(* IEC 61131-3 sources: Codesys_IAP/Demo/PLC1/PLC 1 Simulatie Ladder StructuredTekst IOStructures 2V0_tekst/Programma Structured Text/Structures, 7 files *)

(* ---- hmiIO.st ---- *)
(*#### DECLARATIE ####*)
// Datum : 17 december 2020, Auteur: Gerard Harkema
TYPE hmiIO :
STRUCT
	// Indrukken resetknop
	Ix_Resetknop			: REFERENCE TO BOOL;
	// Keuzeknop staat op hand
	Ix_Hand					: REFERENCE TO BOOL;
	// Keuzeknop staat op auto
	Ix_Auto					: REFERENCE TO BOOL;
	// Indrukken noodstop
	Ix_Noodstop				: REFERENCE TO BOOL;
	// Bekers magazijn zijn op

	// Indrukken startknop
	Ix_Stopknop				: REFERENCE TO BOOL;
	// Indrukken stopknop
	Ix_Startknop			: REFERENCE TO BOOL;
	//Perslucht is aanwezig

	// Visualisatie invisible Gele vlak
	Qx_GeleLamp				: REFERENCE TO BOOL;
	// Visualisatie invisible groene vlak
	Qx_GroeneLamp			: REFERENCE TO BOOL;
	// Visualisatie invisible rode vlak
	Qx_RodeLamp				: REFERENCE TO BOOL;

END_STRUCT
END_TYPE

(* ---- magazijnIO.st ---- *)
(*#### DECLARATIE ####*)
// Datum : 17 december 2020, Auteur: Gerard Harkema
TYPE magazijnIO :
STRUCT
	// Bekers magazijn zijn op
	Ix_MagazijnLeeg				: REFERENCE TO BOOL;
	// Beker is uit dekselmagazijn gestoten
	Ix_UitstoterBekerIn			: REFERENCE TO BOOL;
	// Uitstoter Beker haalt nieuwe beker op
	Ix_UitstoterBekerUit		: REFERENCE TO BOOL;
	// Beker uit magazijn stoten
	Qx_BekerUitstoten			: REFERENCE TO BOOL;

	//Perslucht is aanwezig
	Ix_PersluchtAanwezig 		: REFERENCE TO BOOL;

END_STRUCT
END_TYPE

(* ---- meetstationIO.st ---- *)
(*#### DECLARATIE ####*)
// Datum : 17 december 2020, Auteur: Gerard Harkema
TYPE meetstationIO :
STRUCT
	//Beker aanwezig op detectiepositie
	Ix_BekerAanwezig :REFERENCE TO BOOL;
	//Beker is van aluminium
	Ix_BekerMetaal :REFERENCE TO BOOL;
	//Beker reflecteert en is dus niet zwart
	Ix_BekerReflecteerd :REFERENCE TO BOOL;
END_STRUCT
END_TYPE

(* ---- overzetterIO.st ---- *)
(*#### DECLARATIE ####*)
// Datum : 17 december 2020, Auteur: Gerard Harkema
TYPE overzetterIO :
STRUCT
	//Werkstuk door overzetter opgepakt
	Ix_VacuumAanwezig 		:REFERENCE TO BOOL;
	//Overzetter haalt beker op(linker pos.)
	Ix_OverzetterIsLinks 	:REFERENCE TO BOOL;
	//Overzetter plaatst beker op sorteerpositie
	Ix_OverzetterIsRechts 	:REFERENCE TO BOOL;
	//Beker aanwezig op detectiepositie

		//Beker oppakken
	Qx_VacuumAan 			:REFERENCE TO BOOL;
	//Beker loslaten
	Qx_BekerLossen 			:REFERENCE TO BOOL;
	//Overzetter naar bekermagazijn
	Qx_OverzetterLinks 		:REFERENCE TO BOOL;
	//Overzetter naar sorteerpositie
	Qx_OverzetterRechts 	:REFERENCE TO BOOL;

END_STRUCT
END_TYPE

(* ---- sorteerGootIO.st ---- *)
(*#### DECLARATIE ####*)
// Datum : 17 december 2020, Auteur: Gerard Harkema
TYPE sorteerGootIO :
STRUCT
		//Product is naar een van de goten gegaan
	Ix_BekerInGoot 			:REFERENCE TO BOOL;
	//Pusher uitvoergoot 1 is in
	Ix_UitvoerGoot1IsIn 	:REFERENCE TO BOOL;
	//Pusher uitvoergoot 2 is in
	Ix_UitvoerGoot2IsIn 	:REFERENCE TO BOOL;
	//Pusher uitvoergoot 3 is in
	Ix_UitvoerGoot3IsIn 	:REFERENCE TO BOOL;
	//Beker afvoeren is bezig
	Ix_StationAfvoerVrij 	:REFERENCE TO BOOL;
	//Pusher uitvoergoot 1 is uit
	Ix_UitvoerGoot1IsUit 	:REFERENCE TO BOOL;
	//Pusher uitvoergoot 2 is uit
	Ix_UitvoerGoot2IsUit 	:REFERENCE TO BOOL;
	//Pusher uitvoergoot 3 is uit
	Ix_UitvoerGoot3IsUit 	:REFERENCE TO BOOL;

	//Transportband aan
	Qx_MotorAfvoerAan 		:REFERENCE TO BOOL;
	//Pusher goot 1 uit
	Qx_UitvoerGoot1Uit 		:REFERENCE TO BOOL;
	//Pusher goot 2 uit
	Qx_UitvoerGoot2Uit 		:REFERENCE TO BOOL;
	//Pusher goot 3 uit
	Qx_UitvoerGoot3Uit 		:REFERENCE TO BOOL;
	//Beker stoppen op band voor detectie
	Qx_StopperUit 			:REFERENCE TO BOOL;
	//Uitsorteren is bezet
	Qx_StationBezet 		:REFERENCE TO BOOL;

	uitvoerGoot1			:uitvoerGootIO;
	uitvoerGoot2			:uitvoerGootIO;
	uitvoerGoot3			:uitvoerGootIO;
	meetstation				:meetstationIO;

END_STRUCT
END_TYPE

(* ---- sorteerStationIO.st ---- *)
(*#### DECLARATIE ####*)
// Datum : 17 december 2020, Auteur: Gerard Harkema
TYPE sorteerStationIO :
STRUCT
	magazijn		: magazijnIO;
	overzetter		: overzetterIO;
	sorteerGoot		: sorteerGootIO;
	hmi				: hmiIO;
END_STRUCT
END_TYPE

(* ---- uitvoerGootIO.st ---- *)
(*#### DECLARATIE ####*)
// Datum : 17 december 2020, Auteur: Gerard Harkema
TYPE uitvoerGootIO :
STRUCT
	//Pusher uitvoergoo is in
	Ix_UitvoerGootIsIn 		: REFERENCE TO BOOL;
	//Pusher uitvoergoot is uit
	Ix_UitvoerGootIsUit 	: REFERENCE TO BOOL;
	//Pusher goot uit
	Qx_UitvoerGootUit 		: REFERENCE TO BOOL;
END_STRUCT
END_TYPE
